FUNCTION_BLOCK Controle_Gradeamento_HMI (* Service Interface Function Block Type *)
  (* Standard: 61499-2 *)
  (* Version 1.0, 21/10/2026, Hidryco, Hidryco, IHM do Controle_Gradeamento *)
  PACKAGE Hidryco.HidrycoLib;
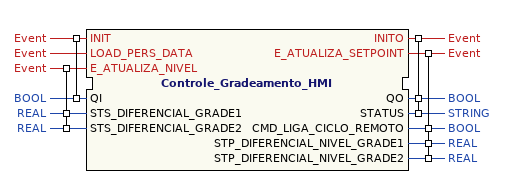
  EVENT_INPUT
    INIT WITH QI;
    LOAD_PERS_DATA; (* Reenvia os parametros persistentes *)
    E_ATUALIZA_NIVEL WITH STS_DIFERENCIAL_GRADE1, STS_DIFERENCIAL_GRADE2; (* Status do processo *)
  END_EVENT
  EVENT_OUTPUT
    INITO WITH QO, STATUS;
    E_ATUALIZA_SETPOINT WITH CMD_LIGA_CICLO_REMOTO, STP_DIFERENCIAL_NIVEL_GRADE1, STP_DIFERENCIAL_NIVEL_GRADE2; (* Ajustes (IHM/OPC UA e LOAD_PERS_DATA) *)
  END_EVENT
  VAR_INPUT
    QI : BOOL;
    STS_DIFERENCIAL_GRADE1 : REAL; (* Nivel diferencial da grade 1 agora (%) *)
    STS_DIFERENCIAL_GRADE2 : REAL; (* Nivel diferencial da grade 2 agora (%) *)
  END_VAR
  VAR_OUTPUT
    QO : BOOL; (* Event Output Qualifier *)
    STATUS : STRING; (* Service Status *)
    CMD_LIGA_CICLO_REMOTO : BOOL; (* Ciclo remoto *)
    STP_DIFERENCIAL_NIVEL_GRADE1 : REAL; (* Diferencial de nível para limpar a grade 1 *)
    STP_DIFERENCIAL_NIVEL_GRADE2 : REAL; (* Diferencial de nível para limpar a grade 2 *)
  END_VAR
  SERVICE /
    SEQUENCE 
    END_SEQUENCE
  END_SERVICE
END_FUNCTION_BLOCK
